{attribute 'qualified_only'}
{attribute 'strict'}
{attribute 'to_string'}
TYPE E_PolarIIChamber_ServiceId :
(
	Chamber_SetMode := 1,
	Chamber_Initial := 2,
	Chamber_SingleProcess := 3,
	Chamber_EMGS := 4,
	Chamber_SetConfig := 5,
	Chamber_ArmAlignTest := 6,
	Chamber_ArmTest := 7,
	Chamber_FlowCalibration := 8,
	Chamber_CupChamberClean := 9,
	Chamber_DoNozzleClean := 10,
	Chamber_DoNozzlePreflush := 11,
	
	Arm1_Lift_TopPos := 1001,
	Arm1_Lift_DownPos := 1002,
	Arm1_Rotate_JogPositive := 1003,
	Arm1_Rotate_JogNegative := 1004,
	Arm1_Rotate_IncrementalJog := 1005,
	Arm1_Rotate_MoveRecipe := 1006,
	Arm1_Rotate_NegLimitPos := 1007,
	Arm1_Rotate_PosLimitPos := 1008,
	Arm1_Rotate_NozPortPos := 1009,
	Arm1_Rotate_Noz1CenterPos := 1010,
	Arm1_Rotate_Noz2CenterPos := 1011,
	Arm1_Rotate_Noz3CenterPos := 1012,
	Arm1_Noz1_ChemicalSupply := 1013,
	Arm1_Noz2_ChemicalSupply := 1014,
	Arm1_Noz3_ChemicalSupply := 1015,
	Arm1_NozPortNoz1_Supply := 1016,
	Arm1_NozPortNoz2_Supply := 1017,
	Arm1_NozPortNoz3_Supply := 1018,
	Arm1_NozPortDrainer_Select1 := 1019,
	Arm1_NozPortDrainer_Select2 := 1020,
	Arm1_NozPortDrainer_Select3 := 1021,
	
	Arm2_Lift_TopPos := 1101,
	Arm2_Lift_DownPos := 1102,
	Arm2_Rotate_JogPositive := 1103,
	Arm2_Rotate_JogNegative := 1104,
	Arm2_Rotate_IncrementalJog := 1105,
	Arm2_Rotate_MoveRecipe := 1106,
	Arm2_Rotate_NegLimitPos := 1107,
	Arm2_Rotate_PosLimitPos := 1108,
	Arm2_Rotate_NozPortPos := 1109,
	Arm2_Rotate_Noz1CenterPos := 1110,
	Arm2_Rotate_Noz2CenterPos := 1111,
	Arm2_Rotate_Noz3CenterPos := 1112,
	Arm2_Noz1_ChemicalSupply := 1113,
	Arm2_Noz2_ChemicalSupply := 1114,
	Arm2_Noz3_ChemicalSupply := 1115,
	Arm2_NozPortNoz1_Supply := 1116,
	Arm2_NozPortNoz2_Supply := 1117,
	Arm2_NozPortNoz3_Supply := 1118,
	Arm2_NozPortDrainer_Select1 := 1119,
	Arm2_NozPortDrainer_Select2 := 1120,
	Arm2_NozPortDrainer_Select3 := 1121,
	
	Arm3_Lift_TopPos := 1201,
	Arm3_Lift_DownPos := 1202,
	Arm3_Rotate_JogPositive := 1203,
	Arm3_Rotate_JogNegative := 1204,
	Arm3_Rotate_IncrementalJog := 1205,
	Arm3_Rotate_MoveRecipe := 1206,
	Arm3_Rotate_NegLimitPos := 1207,
	Arm3_Rotate_PosLimitPos := 1208,
	Arm3_Rotate_Noz1CenterPos := 1209,
	Arm3_Rotate_Noz2CenterPos := 1210,
	Arm3_Noz1_ChemicalSupply := 1211,
	Arm3_Noz2_ChemicalSupply := 1212,

	Arm4_Lift_TopPos := 1301,
	Arm4_Lift_DownPos := 1302,
	Arm4_Rotate_JogPositive := 1303,
	Arm4_Rotate_JogNegative := 1304,
	Arm4_Rotate_IncrementalJog := 1305,
	Arm4_Rotate_MoveRecipe := 1306,
	Arm4_Rotate_NegLimitPos := 1307,
	Arm4_Rotate_PosLimitPos := 1308,
	Arm4_Rotate_Noz1CenterPos := 1309,
	Arm4_Noz1_ChemicalSupply := 1310,
	
	Cup1_Lift_JogPositive := 2001,
	Cup1_Lift_JogNegative := 2002,
	Cup1_Lift_IncrementalJog := 2003,
	Cup1_Lift_DecoupleStop := 2004,
	Cup1_Lift_TopPos := 2005,
	Cup1_Lift_MiddlePos := 2006,
	Cup1_Lift_DownPos := 2007,
	Cup1_Drainer_Select1 := 2008,
	Cup1_Drainer_Select2 := 2009,
	Cup1_Drainer_Select3 := 2010,
	
	Cup2_Lift_JogPositive := 2101,
	Cup2_Lift_JogNegative := 2102,
	Cup2_Lift_IncrementalJog := 2103,
	Cup2_Lift_DecoupleStop := 2104,
	Cup2_Lift_TopPos := 2105,
	Cup2_Lift_MiddlePos := 2106,
	Cup2_Lift_DownPos := 2107,
	Cup2_Drainer_Select1 := 2108,
	Cup2_Drainer_Select2 := 2109,
	Cup2_Drainer_Select3 := 2110,
	
	Cup3_Lift_JogPositive := 2201,
	Cup3_Lift_JogNegative := 2202,
	Cup3_Lift_IncrementalJog := 2203,
	Cup3_Lift_DecoupleStop := 2204,
	Cup3_Lift_TopPos := 2205,
	Cup3_Lift_MiddlePos := 2206,
	Cup3_Lift_DownPos := 2207,
	Cup3_Drainer_Select1 := 2208,
	Cup3_Drainer_Select2 := 2209,
	Cup3_Drainer_Select3 := 2210,
	
	Cup4_Lift_JogPositive := 2301,
	Cup4_Lift_JogNegative := 2302,
	Cup4_Lift_IncrementalJog := 2303,
	Cup4_Lift_DecoupleStop := 2304,
	Cup4_Lift_TopPos := 2305,
	Cup4_Lift_MiddlePos := 2306,
	Cup4_Lift_DownPos := 2307,
	Cup4_Drainer_Select1 := 2308,
	Cup4_Drainer_Select2 := 2309,
	Cup4_Drainer_Select3 := 2310,
	
	Holder_Gripper_Open := 3001,
	Holder_Gripper_Close := 3002,
	Holder_Rotate_OPR := 3003,
	Holder_Rotate_MoveVelocityCW := 3004,
	Holder_Rotate_MoveVelocityCCW := 3005,
	Holder_Rotate_MoveModulo := 3006,
	Holder_VacuumEstablish := 3007,
	
	FixedNoz1_ChemicalSupply := 3101,
	FixedNoz2_ChemicalSupply := 3102,
	FixedNoz3_ChemicalSupply := 3103,
	FixedNoz4_ChemicalSupply := 3104,
	
	OutsideRing_Lift_TopPos := 3201,
	OutsideRing_Lift_DownPos := 3202,
	OutsideRing_Rotate_MoveVelocityCW := 3203,
	OutsideRing_Rotate_MoveVelocityCCW := 3204,
	
	Shutter_Open := 3301,
	Shutter_Close := 3302,
	
	ExhaustFan1_SupplyFlowPID := 3401,
	ExhaustFan2_SupplyFlowPID := 3402,
	ExhaustFan3_SupplyFlowPID := 3403,
	ExhaustFan4_SupplyFlowPID := 3404,
	ExhaustDamper_AEX := 3411,
	ExhaustDamper_SEX := 3412,
	
	SideVent1_Open := 3501,
	SideVent1_Close := 3502,
	SideVent2_Open := 3503,
	SideVent2_Close := 3504,
	SideVent3_Open := 3505,
	SideVent3_Close := 3506,
	SideVent4_Open := 3507,
	SideVent4_Close := 3508
) UDINT;
END_TYPE

(* stored: Version 1.1.0.1, ProductVersion 3.1.4026.18
   DUT E_PolarIIChamber_ServiceId: Id {14000000-0000-0000-0000-000000000001} *)
